Fanuc KAREL source: KT00654.KL

PROGRAM KT00654
%NOLOCKGROUP
VAR
  P1: POSITION
  P2: POSITION
  OUT: BOOLEAN
BEGIN
  OUT = NOT P1
END KT00654
